Fanuc KAREL source: KA00035.KL

PROGRAM KA00035
%NOLOCKGROUP
VAR
  SRC: BOOLEAN
  DST: ARRAY[2] OF BYTE
BEGIN
  SRC = TRUE
  DST[1] = SRC
END KA00035
